{attribute 'qualified_only'}
{attribute 'strict'}
{attribute 'to_string'}
// Run Mode direction / single-end animation location, subindex 10
// (219132 Rev. A, section 1.3.2).
TYPE E_BannerWLS15Pro_Direction :
(
    eUp   := 0,
    eDown := 1
) BYTE;
END_TYPE

(* stored: Version 1.1.0.1
   DUT E_BannerWLS15Pro_Direction: Id {d18b84b4-348e-46ea-8e29-d6a1f18d0502} *)
